// TIA Portal V19 export
VAR_GLOBAL   // PLC tag table "R3_OUT"
   "ByteOUT :0 R3" AT %QB142 : Byte;   // System Bits 1
   "ByteOUT :1 R3" AT %QB143 : Byte;   // System Bits 2
   "ByteOUT :2 R3" AT %QB144 : Byte;   // Signals
   "ByteOUT :3 R3" AT %QB145 : Byte;   // Signals
   "ByteOUT :4 R3" AT %QB146 : Byte;   // CMD
   "ByteOUT :5 R3" AT %QB147 : Byte;   // CMD
   "ByteOUT :6 R3" AT %QB148 : Byte;   // X
   "ByteOUT :7 R3" AT %QB149 : Byte;   // X
   "ByteOUT :8 R3" AT %QB150 : Byte;   // Y
   "ByteOUT :9 R3" AT %QB151 : Byte;   // Y
   "ByteOUT :10 R3" AT %QB152 : Byte;   // Z
   "ByteOUT :11 R3" AT %QB153 : Byte;   // Z
   "ByteOUT :12 R3" AT %QB154 : Byte;
   "ByteOUT :13 R3" AT %QB155 : Byte;
   "ByteOUT :14 R3" AT %QB156 : Byte;
   "ByteOUT :15 R3" AT %QB157 : Byte;
   "ByteOUT :16 R3" AT %QB158 : Byte;
   "ByteOUT :17 R3" AT %QB159 : Byte;
   "ByteOUT :18 R3" AT %QB160 : Byte;
   "ByteOUT :19 R3" AT %QB161 : Byte;
   "ByteOUT :20 R3" AT %QB162 : Byte;
   "ByteOUT :21 R3" AT %QB163 : Byte;
   "ByteOUT :22 R3" AT %QB164 : Byte;
   "ByteOUT :23 R3" AT %QB165 : Byte;
   "ByteOUT :24 R3" AT %QB166 : Byte;
   "ByteOUT :25 R3" AT %QB167 : Byte;
   "ByteOUT :26 R3" AT %QB168 : Byte;
   "ByteOUT :27 R3" AT %QB169 : Byte;
   "ByteOUT :28 R3" AT %QB170 : Byte;
   "ByteOUT :29 R3" AT %QB171 : Byte;
   "ByteOUT :30 R3" AT %QB172 : Byte;
   "ByteOUT :31 R3" AT %QB173 : Byte;
   "ByteOUT :32 R3" AT %QB174 : Byte;
   "ByteOUT :33 R3" AT %QB175 : Byte;
   "ByteOUT :34 R3" AT %QB176 : Byte;
   "ByteOUT :35 R3" AT %QB177 : Byte;
   "ByteOUT :36 R3" AT %QB178 : Byte;
   "ByteOUT :37 R3" AT %QB179 : Byte;
   "ByteOUT :38 R3" AT %QB180 : Byte;
   "ByteOUT :39 R3" AT %QB181 : Byte;
   "ByteOUT :40 R3" AT %QB182 : Byte;
   "ByteOUT :41 R3" AT %QB183 : Byte;
   "ByteOUT :42 R3" AT %QB184 : Byte;
   "ByteOUT :43 R3" AT %QB185 : Byte;
   "ByteOUT :44 R3" AT %QB186 : Byte;
   "ByteOUT :45 R3" AT %QB187 : Byte;
   "ByteOUT :46 R3" AT %QB188 : Byte;
   "ByteOUT :47 R3" AT %QB189 : Byte;
   "ByteOUT :48 R3" AT %QB190 : Byte;
   "ByteOUT :49 R3" AT %QB191 : Byte;
   "ByteOUT :50 R3" AT %QB192 : Byte;
   "ByteOUT :51 R3" AT %QB193 : Byte;
   "ByteOUT :52 R3" AT %QB194 : Byte;
   "ByteOUT :53 R3" AT %QB195 : Byte;
   "ByteOUT :54 R3" AT %QB196 : Byte;
   "ByteOUT :55 R3" AT %QB197 : Byte;
   "ByteOUT :56 R3" AT %QB198 : Byte;
   "ByteOUT :57 R3" AT %QB199 : Byte;
   "ByteOUT :58 R3" AT %QB200 : Byte;
   "ByteOUT :59 R3" AT %QB201 : Byte;
   "ByteOUT :60 R3" AT %QB202 : Byte;
   "ByteOUT :61 R3" AT %QB203 : Byte;
   "ByteOUT :62 R3" AT %QB204 : Byte;
   "ByteOUT :63 R3" AT %QB205 : Byte;
END_VAR
